(* IEC 61131-3 sources: llm-plc-st-eval/data/processed_definitivo/claude-sonnet-4-6/I5/few_shot, 3 files *)

(* ---- ejec_1.st ---- *)
FUNCTION_BLOCK FB_Clasificadora
VAR_INPUT
    sensorPresencia : BOOL; (* Sensor de paso de pieza *)
    sensorAltura    : BOOL; (* Sensor de pieza alta *)
END_VAR
VAR_OUTPUT
    banda   : BOOL; (* Banda transportadora activa *)
    piston  : BOOL; (* Piston desviador *)
    nAltas  : INT;  (* Contador de piezas altas *)
    nBajas  : INT;  (* Contador de piezas bajas *)
END_VAR
VAR
    tRetardo : TON; (* Temporizador de retardo 2 s hasta el desviador *)
    tPulso   : TP;  (* Temporizador de pulso 1 s del piston *)
    rPresencia : R_TRIG; (* Flanco ascendente del sensor de presencia *)
    piezaAlta  : BOOL;   (* Indica que la pieza detectada es alta *)
END_VAR

(* La banda funciona continuamente *)
banda := TRUE;

(* Detectar flanco ascendente del sensor de presencia *)
rPresencia(CLK := sensorPresencia);

IF rPresencia.Q THEN
    IF sensorAltura THEN
        (* Pieza alta: registrar y armar retardo *)
        nAltas    := nAltas + 1;
        piezaAlta := TRUE;
    ELSE
        (* Pieza baja: solo registrar *)
        nBajas := nBajas + 1;
    END_IF;
END_IF;

(* Retardo de 2 s: la pieza tarda ese tiempo en llegar al desviador *)
tRetardo(IN := piezaAlta, PT := T#2S);

(* Al cumplirse el retardo, lanzar pulso de 1 s en el piston *)
tPulso(IN := tRetardo.Q, PT := T#1S);

(* Cuando el pulso termina, desactivar la bandera de pieza alta *)
IF tPulso.Q = FALSE AND tRetardo.Q THEN
    (* El pulso TP.Q cae al terminar; limpiar cuando TP ya no este activo *)
    (* Se limpia piezaAlta cuando el temporizador de pulso finaliza *)
    piezaAlta := FALSE;
END_IF;

(* Activar piston durante el pulso de 1 s *)
piston := tPulso.Q;

END_FUNCTION_BLOCK

(* ---- ejec_2.st ---- *)
FUNCTION_BLOCK FB_Clasificadora
VAR_INPUT
    sensorPresencia : BOOL; (* Sensor de paso de pieza *)
    sensorAltura    : BOOL; (* TRUE = pieza alta *)
END_VAR
VAR_OUTPUT
    banda   : BOOL; (* Banda transportadora activa *)
    piston  : BOOL; (* Pistón desviador *)
    nAltas  : INT;  (* Contador de piezas altas *)
    nBajas  : INT;  (* Contador de piezas bajas *)
END_VAR
VAR
    rPresencia  : R_TRIG; (* Flanco ascendente de sensorPresencia *)
    tRetardo    : TON;    (* Retardo de 2 s hasta el desviador *)
    tPulso      : TP;     (* Pulso de 1 s del pistón *)
    bEsAlta     : BOOL;   (* Indica que la pieza detectada es alta *)
END_VAR

(* La banda funciona siempre *)
banda := TRUE;

(* Detectar flanco ascendente de presencia de pieza *)
rPresencia(CLK := sensorPresencia);

IF rPresencia.Q THEN
    IF sensorAltura THEN
        (* Pieza alta: registrar y armar retardo *)
        nAltas  := nAltas + 1;
        bEsAlta := TRUE;
    ELSE
        (* Pieza baja: solo contar *)
        nBajas  := nBajas + 1;
        bEsAlta := FALSE;
    END_IF;
END_IF;

(* Retardo de 2 s: arranca cuando hay pieza alta pendiente *)
tRetardo(IN := bEsAlta, PT := T#2S);

(* Al cumplirse el retardo, disparar el pulso del pistón y limpiar la bandera *)
IF tRetardo.Q THEN
    bEsAlta := FALSE; (* Evita rearrancar el retardo *)
END_IF;

(* Pulso de 1 s del pistón, iniciado por el flanco de salida del retardo *)
tPulso(IN := tRetardo.Q, PT := T#1S);
piston := tPulso.Q;

END_FUNCTION_BLOCK

(* ---- ejec_3.st ---- *)
FUNCTION_BLOCK FB_Clasificadora
VAR_INPUT
    sensorPresencia : BOOL; (* Sensor de paso de pieza *)
    sensorAltura    : BOOL; (* Sensor de altura: TRUE = pieza alta *)
END_VAR
VAR_OUTPUT
    banda   : BOOL; (* Banda transportadora activa *)
    piston  : BOOL; (* Pistón desviador *)
    nAltas  : INT;  (* Contador de piezas altas *)
    nBajas  : INT;  (* Contador de piezas bajas *)
END_VAR
VAR
    tRetardo : TON; (* Retardo de 2 s hasta llegar al desviador *)
    tPulso   : TP;  (* Pulso de 1 s para activar el pistón *)
    rPresencia : R_TRIG; (* Flanco ascendente del sensor de presencia *)
    bPiezaAlta : BOOL;   (* Indica que la pieza detectada es alta *)
END_VAR

(* La banda funciona siempre *)
banda := TRUE;

(* Detectar flanco ascendente del sensor de presencia *)
rPresencia(CLK := sensorPresencia);

IF rPresencia.Q THEN
    IF sensorAltura THEN
        (* Pieza alta: registrar y armar retardo *)
        nAltas     := nAltas + 1;
        bPiezaAlta := TRUE;
    ELSE
        (* Pieza baja: solo contar *)
        nBajas := nBajas + 1;
    END_IF;
END_IF;

(* Retardo de 2 s: la pieza tarda ese tiempo en llegar al desviador *)
tRetardo(IN := bPiezaAlta, PT := T#2S);

(* Al cumplirse el retardo, lanzar pulso de 1 s en el pistón *)
tPulso(IN := tRetardo.Q, PT := T#1S);

(* Cuando el pulso termina, limpiar la bandera de pieza alta *)
IF NOT tPulso.Q AND NOT tRetardo.Q AND bPiezaAlta THEN
    (* El temporizador de retardo aún no ha arrancado o ya terminó el pulso *)
    (* Limpiar solo cuando el ciclo completo haya concluido *)
    IF tRetardo.ET = T#0S AND NOT tRetardo.IN THEN
        bPiezaAlta := FALSE;
    END_IF;
END_IF;

(* Limpiar bandera al finalizar el pulso del pistón *)
IF tPulso.Q = FALSE AND tRetardo.Q = FALSE AND tRetardo.ET >= T#2S THEN
    bPiezaAlta := FALSE;
END_IF;

(* Activar pistón durante el pulso de 1 s *)
piston := tPulso.Q;

END_FUNCTION_BLOCK
